// TIA Portal V20 export
Screen "Main"  1276x673
  ScreenItem "permanentareaborderrectangle" at 0,0 size 0x0  Type=HmiRectangle
  ScreenItem "Overview_01_Shadow_3" at 5,6 size 217x208  Type=HmiRectangle
  ScreenItem "Overview_1" at 0,0 size 217x208  Type=HmiRectangle
  ScreenItem "PosDev_Lifter_3" at 5,73 size 207x125  Type=HmiGraphicView
  ScreenItem "Overview_01_Text_3" at 2,4 size 212x31  Type=HmiTextBox
  ScreenItem "Overview_01_TextTyp_3" at 2,38 size 180x26  Type=HmiTextBox
  ScreenItem "Overview_01_Button_1" at 2,4 size 217x208  Type=HmiButton
  ScreenItem "Overview_01_Button_6" at 2,4 size 217x208  Type=HmiButton
  ScreenItem "Overview_01_Shadow_1" at 5,6 size 217x208  Type=HmiRectangle
  ScreenItem "Overview_2" at 0,0 size 217x208  Type=HmiRectangle
  ScreenItem "PosDev_Lifter_1" at 5,73 size 207x125  Type=HmiGraphicView
  ScreenItem "Overview_01_Text_1" at 2,4 size 212x31  Type=HmiTextBox
  ScreenItem "Overview_01_TextTyp_1" at 2,38 size 180x26  Type=HmiTextBox
  ScreenItem "Overview_01_Button_2" at 1,1 size 217x208  Type=HmiButton
  ScreenItem "Overview_01_Button_3" at 1,3 size 217x208  Type=HmiButton
  ScreenItem "Overview_01_Shadow_4" at 5,6 size 217x208  Type=HmiRectangle
  ScreenItem "Overview_4" at 0,0 size 217x208  Type=HmiRectangle
  ScreenItem "PosDev_Lifter_4" at 5,73 size 207x125  Type=HmiGraphicView
  ScreenItem "Overview_01_Text_4" at 2,4 size 212x31  Type=HmiTextBox
  ScreenItem "Overview_01_TextTyp_4" at 2,38 size 180x26  Type=HmiTextBox
  ScreenItem "Overview_01_Button_7" at 1,3 size 217x208  Type=HmiButton
  ScreenItem "Overview_01_Button_8" at 1,2 size 217x208  Type=HmiButton
  ScreenItem "Overview_01_Shadow_2" at 5,6 size 217x208  Type=HmiRectangle
  ScreenItem "Overview_3" at 0,0 size 217x208  Type=HmiRectangle
  ScreenItem "PosDev_Lifter_2" at 5,73 size 207x125  Type=HmiGraphicView
  ScreenItem "Overview_01_Text_2" at 2,4 size 212x31  Type=HmiTextBox
  ScreenItem "Overview_01_TextTyp_2" at 2,38 size 180x26  Type=HmiTextBox
  ScreenItem "Overview_01_Button_4" at 2,3 size 217x208  Type=HmiButton
  ScreenItem "Overview_01_Button_5" at 2,3 size 217x208  Type=HmiButton
